// TIA Portal V21 export
// export: Created 2026-11-10T07:35:08.2891503Z, ExportSetting WithDefaults, DisplayName Totally Integrated Automation Portal, DisplayVersion V21 Update 3, DisplayName STEP 7 Professional, DisplayVersion V21 Update 3, DisplayName STEP 7 Safety, DisplayVersion V21, DisplayName Tech WebApplication, DisplayVersion V21, DisplayName WinCC Basic/Comfort/Advanced, DisplayVersion V21 Update 3, DisplayName WinCC Unified, DisplayVersion V21 Update 3
FUNCTION_BLOCK "FB_Lad_ex064"   // FB22, LAD
{ S7_Optimized_Access := 'TRUE' }
VERSION : 0.1
// stored: AutoNumber true, IsIECCheckEnabled false, IsRetainMemResEnabled false, MemoryReserve 100, SetENOAutomatically false, UDAEnableTagReadback false
   VAR_INPUT
      v_req : Bool;
      v_laddr : HW_INTERFACE;
      v_group : Byte;
      v_mode : Byte;
      v_ret_val : Int;
   END_VAR
   VAR_OUTPUT
      v_busy : Bool;
   END_VAR
BEGIN

REGION Network 1: DPSYC_FR - Synchronize DP slaves / Freeze inputs
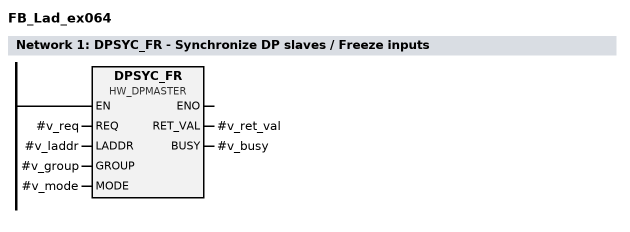
   RUNG wire#powerrail
      { S7_Templates := "laddr_type := HW_DPMASTER" } DPSYC_FR(REQ := #v_req, LADDR := #v_laddr, GROUP := #v_group, MODE := #v_mode, RET_VAL => #v_ret_val, BUSY => #v_busy)
   END_RUNG
   // the same network as SCL:
   #v_ret_val := DPSYC_FR(REQ := #v_req, LADDR := #v_laddr, GROUP := #v_group, MODE := #v_mode, BUSY => #v_busy);
END_REGION
END_FUNCTION_BLOCK
